(*
Citation references, like [CIT2002]_. Note that citations may get rearranged, e.g., to the bottom of the "page". 

| Some sample text to get some text in between.
| Some sample text to get some text in between.
| Some sample text to get some text in between.
| Some sample text to get some text in between.
| Some sample text to get some text in between.
| Some sample text to get some text in between.

.. [CIT2002] This is the citation.  It's just like a footnote,
   except the label is textual. 

Given a citation like [this]_, one can also refer to it like this_. 

| Some sample text to get some text in between.
| Some sample text to get some text in between.
| Some sample text to get some text in between.
| Some sample text to get some text in between.
| Some sample text to get some text in between.
| Some sample text to get some text in between.

.. [this] here.

| Some sample text to get some text in between.
| Some sample text to get some text in between.
| Some sample text to get some text in between.
| Some sample text to get some text in between.
| Some sample text to get some text in between.
| Some sample text to get some text in between.

*)

FUNCTION_BLOCK FB_Libdoc_Citation
VAR_INPUT
    nVarA : INT;
    nVarB : INT;
END_VAR
VAR_OUTPUT
    nSum : INT;
END_VAR
VAR
END_VAR

END_FUNCTION_BLOCK

(* stored: Version 1.1.0.1, ProductVersion 3.1.4024.0
   POU FB_Libdoc_Citation: Id {73b32be0-ee3b-4855-b606-424fa250e28e}, SpecialFunc None *)
